// TwinCAT 3 PLC project PLC
// ProgramVersion: 3.1.4026.27
// libraries:
//   Tc2_Standard, * (Beckhoff Automation GmbH)
//   Tc2_System, * (Beckhoff Automation GmbH)
//   Tc3_EventLogger, * (Beckhoff Automation GmbH)
// project tree:
//   / PlcTask.TcTTO
//   POUs/ MAIN.TcPOU, FB_ActiveAlarmListener.TcPOU, I_ActiveAlarmList.TcIO, FB_Station.TcPOU, FB_StackLight.TcPOU
//   DUTs/ ST_EventListEntry.TcDUT
//   GVLs/ GVL_Params.TcGVL
// real-time tasks:
//   TASK PlcTask: cycle T#10ms, priority 20, ADS port 350

CONFIGURATION PLC
    RESOURCE PLC ON TwinCAT3
        TASK PlcTask(INTERVAL := T#10ms, PRIORITY := 20);
        PROGRAM MAIN WITH PlcTask : MAIN;
    END_RESOURCE
END_CONFIGURATION

// ---- DUTs/ST_EventListEntry.TcDUT
// One row of FB_ActiveAlarmListener (active alarm table and message ring buffer).
// Application independent: everything FB_TcEvent exposes, copied out of the callback.
TYPE ST_EventListEntry :
STRUCT
    bUsed       : BOOL;             // row in use = alarm is ACTIVE (raised, or cleared but waiting for confirmation)
    bIsAlarm    : BOOL;             // TRUE = alarm, FALSE = message
    bRaised     : BOOL;             // alarm state: TRUE = Raised, FALSE = cleared (row only kept while waiting for confirmation)
    eConfirmationState : TcEventConfirmationState;  // NotSupported / NotRequired / WaitForConfirmation / Confirmed / Reset
    nSequence   : UDINT;            // running number (messages only)
    eventClass  : GUID;             // event class
    nEventId    : UDINT;            // event id within the class
    eSeverity   : TcEventSeverity;  // Verbose..Critical
    nTimestamp  : ULINT;            // raise / send time stamped by the EventLogger, 100 ns since 1601-01-01 UTC
    nReceived   : ULINT;            // F_GetSystemTime when the listener callback ran (same clock, same unit)
    tLatency    : LTIME;            // nReceived - nTimestamp: raise -> visible in this table
    nSourceId   : UDINT;            // I_TcSourceInfo.nId   (application defined, e.g. station number)
    guidSource  : GUID;             // I_TcSourceInfo.guid
    sSourceName : STRING(255);      // I_TcSourceInfo.sName
END_STRUCT
END_TYPE

// ---- GVLs/GVL_Params.TcGVL
// Application (test harness) parameters.
{attribute 'qualified_only'}
VAR_GLOBAL CONSTANT
    cStations        : UDINT := 12;      // number of stations / stack lights
    cStationAlarms   : UDINT := 8;       // alarms per station (FB_Station.aAlarms, Event3..Event10)
END_VAR

// ---- POUs/I_ActiveAlarmList.TcIO
// Read-only view of an "active alarm list" + recent-message ring buffer.
//
// Consumers (stack lights, HMI summaries, interlocks, ...) depend on THIS, not on the
// FB that produces the list. FB_ActiveAlarmListener implements it from EventLogger
// callbacks; any other producer (e.g. a list built from the PLC's own FB_TcAlarm.bRaised
// states, or one fed by the .NET proxy over ADS) can implement it too and the consumers
// do not change.
//
// Alarm identity = event class + event id + source id.
// Rows are addressed 1..nMaxAlarms; GetAlarm is FALSE for an empty row.
// Messages are addressed by running sequence number 1..nMessageSequence; GetMessage is
// FALSE once a message has been overwritten in the ring buffer (size nMaxRecentMessages).
INTERFACE I_ActiveAlarmList EXTENDS __SYSTEM.IQueryInterface

// Number of raised alarms (any source) whose severity is within [eMinSeverity .. eMaxSeverity].
METHOD Count : UDINT
VAR_INPUT
    eMinSeverity : TcEventSeverity;
    eMaxSeverity : TcEventSeverity;
END_VAR
END_METHOD

// Number of raised alarms from source nSourceId (= FB_TcSourceInfo.nId the publisher used)
// whose severity is within [eMinSeverity .. eMaxSeverity].
METHOD CountBySource : UDINT
VAR_INPUT
    nSourceId    : UDINT;
    eMinSeverity : TcEventSeverity;
    eMaxSeverity : TcEventSeverity;
END_VAR
END_METHOD

// Number of raised alarms of one event class whose severity is within [eMinSeverity .. eMaxSeverity].
METHOD CountByEventClass : UDINT
VAR_INPUT
    eventClass   : GUID;
    eMinSeverity : TcEventSeverity;
    eMaxSeverity : TcEventSeverity;
END_VAR
END_METHOD

// TRUE if the alarm (event class + event id + source id) is currently raised.
METHOD IsActive : BOOL
VAR_INPUT
    eventClass : GUID;
    nEventId   : UDINT;
    nSourceId  : UDINT;
END_VAR
END_METHOD

// Copies row nIndex (1..nMaxAlarms) of the active alarm table. FALSE if the row is empty
// or nIndex is out of range. Iterate 1..nMaxAlarms to enumerate all raised alarms.
METHOD GetAlarm : BOOL
VAR_INPUT
    nIndex : UDINT;
END_VAR
VAR_IN_OUT
    stEntry : ST_EventListEntry;
END_VAR
END_METHOD

// Fetches the message with running number nSequence from the ring buffer.
// Returns FALSE if that message was never received or has already been overwritten.
// Typical use: remember nMessageSequence, then loop over the newer ones each cycle.
METHOD GetMessage : BOOL
VAR_INPUT
    nSequence : UDINT;
END_VAR
VAR_IN_OUT
    stEntry : ST_EventListEntry;
END_VAR
END_METHOD

// Number of alarms currently raised (rows in use).
PROPERTY nActiveAlarms : UDINT
GET
END_GET
END_PROPERTY

// Highest valid row index for GetAlarm.
PROPERTY nMaxAlarms : UDINT
GET
END_GET
END_PROPERTY

// Increments on every raise / clear / dispose. Compare to the last value seen to detect "list changed".
PROPERTY nAlarmChangeCounter : UDINT
GET
END_GET
END_PROPERTY

// Running number of the newest message received (0 = none yet).
PROPERTY nMessageSequence : UDINT
GET
END_GET
END_PROPERTY

// Ring buffer size: messages older than nMessageSequence - nMaxRecentMessages are gone.
PROPERTY nMaxRecentMessages : UDINT
GET
END_GET
END_PROPERTY

END_INTERFACE

// ---- POUs/MAIN.TcPOU
// Test harness: 12 stations publish events, ONE listener keeps the active alarm
// list and drives 12 stack lights - all in the PLC, no HMI involved.
//
// How to play (online, in the declaration part of MAIN):
//   1. set nTestStation (1..12) and nTestAlarm (1..8, see FB_Station header for the mapping)
//   2. pulse bTestRaise / bTestClear / bTestSendMessage
//   3. watch aActiveAlarms, aRecentMessages, aStackLights[n].bRed/bYellow/bGreen
PROGRAM MAIN
VAR
    aStations    : ARRAY[1..GVL_Params.cStations] OF FB_Station;      // event publishers (app specific)
    aStackLights : ARRAY[1..GVL_Params.cStations] OF FB_StackLight;   // decoder ring -> outputs (app specific)

    // the generic "active alarm list" (one per PLC) + the storage it works on (sized here, by the application)
    fbListener      : FB_ActiveAlarmListener;
    aActiveAlarms   : ARRAY[1..128] OF ST_EventListEntry;   // raised alarms
    aRecentMessages : ARRAY[1..32]  OF ST_EventListEntry;   // last 32 messages (ring buffer)
    fbFilter        : FB_TcEventFilter;
    bSubscribe   : BOOL := TRUE;
    hrSubscribe  : HRESULT;

    // --- test controls -------------------------------------------------------
    nTestStation       : UDINT := 1;   // 1..12
    nTestAlarm         : UDINT := 1;   // 1..8: 1,4,5 = Warning (yellow)  2,6,7 = Error (red)  3,8 = Critical (red)
    bTestRaise         : BOOL;         // raise aAlarms[nTestAlarm] on station nTestStation
    bTestClear         : BOOL;         // clear it again
    bTestSendMessage   : BOOL;         // green pulse
    bTestClearAll      : BOOL;         // clear every raised alarm on nTestStation
    hrTest             : HRESULT;

    // --- "noise" from another event class, to prove the filter ----------------
    // TC_EVENTS.MachineEvents is NOT in the listener's filter, so these must never
    // show up in fbListener even though they share source id 3 with station 3.
    fbMachineSource    : FB_TcSourceInfo;
    fbMachineMessage   : FB_TcMessage;
    fbMachineAlarm     : FB_TcAlarm;
    bMachineInit       : BOOL := TRUE;
    bTestMachineMessage    : BOOL;
    bTestMachineRaiseAlarm : BOOL;
    bTestMachineClearAlarm : BOOL;
    hrMachineTest      : HRESULT;

    // --- alarm WITH confirmation required: stays in the list after Clear(FALSE) until Confirm(); Clear(TRUE) ends it ---
    fbAckSource        : FB_TcSourceInfo;
    fbAckAlarm         : FB_TcAlarm;            // StationEvents.MotorFault, bWithConfirmation := TRUE, source id 13
    bAckInit           : BOOL := TRUE;
    bTestAckRaise      : BOOL;
    bTestAckConfirm    : BOOL;
    bTestAckClear      : BOOL;                  // Clear(FALSE): confirmation still required
    bTestAckClearReset : BOOL;                  // Clear(TRUE):  confirmation reset
    hrAckTest          : HRESULT;

    i : UDINT;
END_VAR

// 1) stations: give each its id and let it create its events (first cycle)
FOR i := 1 TO GVL_Params.cStations DO
    aStations[i].nStationId := i;
    aStations[i]();
END_FOR

// 2) subscribe the listener once - only to our station event class
IF bSubscribe THEN
    bSubscribe := FALSE;
    // TC_EVENTS.StationEvents is only a namespace; the class GUID is reachable through any of its
    // events (all carry the same uuidEventClass), so this matches ALL events of StationEvents.
    fbFilter.Clear().EventClass.EqualTo(TC_EVENTS.StationEvents.CycleComplete.uuidEventClass);
    hrSubscribe := fbListener.Subscribe2(fbFilter);
END_IF

// 3) process the event queue -> active alarm list (the FB body binds the arrays and runs Execute)
fbListener(aActiveAlarms := aActiveAlarms, aRecentMessages := aRecentMessages);

// 4) stack lights - each one filters the shared list by its own source id.
//    They see the listener only as I_ActiveAlarmList (fbListener is implicitly converted).
FOR i := 1 TO GVL_Params.cStations DO
    aStackLights[i](ipAlarmList := fbListener, nSourceId := i);
END_FOR

// 5) test controls
IF nTestStation >= 1 AND nTestStation <= GVL_Params.cStations THEN
    IF bTestSendMessage THEN bTestSendMessage := FALSE; hrTest := aStations[nTestStation].SendMessage();  END_IF
    IF bTestRaise       THEN bTestRaise       := FALSE; hrTest := aStations[nTestStation].Raise(nTestAlarm); END_IF
    IF bTestClear       THEN bTestClear       := FALSE; hrTest := aStations[nTestStation].Clear(nTestAlarm); END_IF
    IF bTestClearAll    THEN bTestClearAll    := FALSE; aStations[nTestStation].ClearAll();                  END_IF
END_IF

// 6) unrelated event class (filter test)
IF bMachineInit THEN
    bMachineInit := FALSE;
    fbMachineSource.Clear();
    fbMachineSource.nId   := 3;                 // deliberately collides with station 3
    fbMachineSource.sName := 'Machine';
    hrMachineTest := fbMachineMessage.CreateEx(TC_EVENTS.MachineEvents.MachineMessage, fbMachineSource);
    hrMachineTest := fbMachineAlarm.CreateEx(TC_EVENTS.MachineEvents.MachineAlarm, FALSE, fbMachineSource);
END_IF
IF bTestMachineMessage    THEN bTestMachineMessage    := FALSE; hrMachineTest := fbMachineMessage.Send(0);       END_IF
IF bTestMachineRaiseAlarm THEN bTestMachineRaiseAlarm := FALSE; hrMachineTest := fbMachineAlarm.Raise(0);        END_IF
IF bTestMachineClearAlarm THEN bTestMachineClearAlarm := FALSE; hrMachineTest := fbMachineAlarm.Clear(0, FALSE); END_IF

// 7) alarm with confirmation required (source id 13, no stack light; watch aActiveAlarms)
IF bAckInit THEN
    bAckInit := FALSE;
    fbAckSource.Clear();
    fbAckSource.nId   := 13;
    fbAckSource.sName := 'Ack test';
    hrAckTest := fbAckAlarm.CreateEx(TC_EVENTS.StationEvents.MotorFault, TRUE, fbAckSource);
END_IF
IF bTestAckRaise      THEN bTestAckRaise      := FALSE; hrAckTest := fbAckAlarm.Raise(0);        END_IF
IF bTestAckConfirm    THEN bTestAckConfirm    := FALSE; hrAckTest := fbAckAlarm.Confirm(0);      END_IF
IF bTestAckClear      THEN bTestAckClear      := FALSE; hrAckTest := fbAckAlarm.Clear(0, FALSE); END_IF
IF bTestAckClearReset THEN bTestAckClearReset := FALSE; hrAckTest := fbAckAlarm.Clear(0, TRUE);  END_IF

END_PROGRAM

// ---- POUs/FB_Station.TcPOU
// Reusable per-station event publisher.
// All events of a station share one FB_TcSourceInfo whose nId = station number and
// sName = 'Station n'. The listener uses nId to route the event to the right stack light.
//
// Event class TC_EVENTS.StationEvents (MyEvents.tmc), alarm index -> event:
//   message        CycleComplete   Info      'Cycle complete'
//   aAlarms[1]     MaintenanceDue  Warning   'Maintenance due'
//   aAlarms[2]     PartJam         Error     'Part jam'
//   aAlarms[3]     Overtemperature Critical  'Overtemperature'
//   aAlarms[4]     LowMaterial     Warning   'Low material'
//   aAlarms[5]     DoorOpen        Warning   'Door open'
//   aAlarms[6]     MotorFault      Error     'Motor fault'
//   aAlarms[7]     SensorFault     Error     'Sensor fault'
//   aAlarms[8]     EmergencyStop   Critical  'Emergency stop'
// Several alarms share a severity on purpose: the stack light must stay on until the
// LAST raised alarm of that severity is cleared.
FUNCTION_BLOCK FB_Station
VAR_INPUT
    nStationId : UDINT;     // 1..GVL_Params.cStations - set before the first call
END_VAR
VAR_OUTPUT
    bInitialized : BOOL;
    hrLastError  : HRESULT;                                        // last failed call (latched)
    aRaised      : ARRAY[1..GVL_Params.cStationAlarms] OF BOOL;    // live state of this station's own alarms
    nRaised      : UDINT;                                          // how many of them are raised
END_VAR
VAR
    fbSource   : FB_TcSourceInfo;
    fbMessage  : FB_TcMessage;
    aAlarms    : ARRAY[1..GVL_Params.cStationAlarms] OF FB_TcAlarm;
    aAlarmDefs : ARRAY[1..GVL_Params.cStationAlarms] OF TcEventEntry;
    hr         : HRESULT;
    i          : UDINT;
END_VAR

IF NOT bInitialized AND nStationId > 0 THEN
    bInitialized := TRUE;

    // source info = station identity (captured by the events at Create time)
    fbSource.Clear();
    fbSource.nId   := nStationId;
    fbSource.sName := CONCAT('Station ', UDINT_TO_STRING(nStationId));

    aAlarmDefs[1] := TC_EVENTS.StationEvents.MaintenanceDue;
    aAlarmDefs[2] := TC_EVENTS.StationEvents.PartJam;
    aAlarmDefs[3] := TC_EVENTS.StationEvents.Overtemperature;
    aAlarmDefs[4] := TC_EVENTS.StationEvents.LowMaterial;
    aAlarmDefs[5] := TC_EVENTS.StationEvents.DoorOpen;
    aAlarmDefs[6] := TC_EVENTS.StationEvents.MotorFault;
    aAlarmDefs[7] := TC_EVENTS.StationEvents.SensorFault;
    aAlarmDefs[8] := TC_EVENTS.StationEvents.EmergencyStop;

    hr := fbMessage.CreateEx(TC_EVENTS.StationEvents.CycleComplete, fbSource);
    IF FAILED(hr) THEN hrLastError := hr; END_IF
    FOR i := 1 TO GVL_Params.cStationAlarms DO
        hr := aAlarms[i].CreateEx(aAlarmDefs[i], FALSE, fbSource);
        IF FAILED(hr) THEN hrLastError := hr; END_IF
    END_FOR
END_IF

nRaised := 0;
FOR i := 1 TO GVL_Params.cStationAlarms DO
    aRaised[i] := aAlarms[i].bRaised;
    IF aRaised[i] THEN nRaised := nRaised + 1; END_IF
END_FOR

METHOD SendMessage : HRESULT
SendMessage := fbMessage.Send(0);
IF FAILED(SendMessage) THEN hrLastError := SendMessage; END_IF
END_METHOD

// Raises alarm nAlarm (1..GVL_Params.cStationAlarms, see table in the FB header).
METHOD Raise : HRESULT
VAR_INPUT
    nAlarm : UDINT;
END_VAR
IF nAlarm < 1 OR nAlarm > GVL_Params.cStationAlarms THEN
    Raise := DWORD_TO_DINT(16#80070057);  // E_INVALIDARG
ELSE
    Raise := aAlarms[nAlarm].Raise(0);
END_IF
IF FAILED(Raise) THEN hrLastError := Raise; END_IF
END_METHOD

// Clears alarm nAlarm (1..GVL_Params.cStationAlarms).
METHOD Clear : HRESULT
VAR_INPUT
    nAlarm : UDINT;
END_VAR
IF nAlarm < 1 OR nAlarm > GVL_Params.cStationAlarms THEN
    Clear := DWORD_TO_DINT(16#80070057);  // E_INVALIDARG
ELSE
    Clear := aAlarms[nAlarm].Clear(0, FALSE);
END_IF
IF FAILED(Clear) THEN hrLastError := Clear; END_IF
END_METHOD

// Clears every raised alarm of this station (test helper).
METHOD ClearAll
VAR
    n : UDINT;
END_VAR
FOR n := 1 TO GVL_Params.cStationAlarms DO
    IF aAlarms[n].bRaised THEN
        aAlarms[n].Clear(0, FALSE);
    END_IF
END_FOR
END_METHOD

END_FUNCTION_BLOCK

// ---- POUs/FB_StackLight.TcPOU
// APPLICATION SPECIFIC decoder ring: active alarm list -> one station's stack light.
// All knowledge about "stations" lives here; FB_ActiveAlarmListener knows nothing about them.
//   RED    flashes while any Error/Critical alarm from this source is raised
//   YELLOW flashes while any Warning (or lower) alarm from this source is raised
//   GREEN  flashes for 3 s after a message from this source
// The three colors are independent (a stack light can show more than one).
//
// Depends only on I_ActiveAlarmList, not on FB_ActiveAlarmListener: any list producer
// that implements the interface can drive it.
FUNCTION_BLOCK FB_StackLight
VAR_INPUT
    ipAlarmList   : I_ActiveAlarmList;      // the shared list (assign once; 0 = outputs stay off)
    nSourceId     : UDINT;                  // FB_TcSourceInfo.nId this station publishes with
END_VAR
VAR_OUTPUT
    bRed    : BOOL;
    bYellow : BOOL;
    bGreen  : BOOL;
    nActiveAlarms   : UDINT;                // diagnostics
    nActiveWarnings : UDINT;
    bMessageActive  : BOOL;
END_VAR
VAR
    bFirstCycle  : BOOL := TRUE;
    nLastMsgSeq  : UDINT;                   // last message sequence handled
    stMsg        : ST_EventListEntry;
    fbMsgTimer   : TON;
    fbBlinkTimer : TON;
    bBlink       : BOOL;
END_VAR
VAR CONSTANT
    tBlinkHalfPeriod : TIME := T#500MS;     // flash clock (1 Hz)
    tMsgFlashTime    : TIME := T#3S;        // how long GREEN flashes after a message
END_VAR

IF ipAlarmList = 0 THEN                     // no list connected -> everything off
    nActiveAlarms := 0; nActiveWarnings := 0; bMessageActive := FALSE;
    bRed := FALSE; bYellow := FALSE; bGreen := FALSE;
    RETURN;
END_IF

// --- alarms: just count rows of "my" source in the shared list ---
nActiveAlarms   := ipAlarmList.CountBySource(nSourceId, TcEventSeverity.Error,   TcEventSeverity.Critical);
nActiveWarnings := ipAlarmList.CountBySource(nSourceId, TcEventSeverity.Verbose, TcEventSeverity.Warning);

// --- messages: walk the ones that arrived since last cycle, react to "mine" ---
IF bFirstCycle THEN
    bFirstCycle := FALSE;
    nLastMsgSeq := ipAlarmList.nMessageSequence;
END_IF
IF ipAlarmList.nMessageSequence - nLastMsgSeq > ipAlarmList.nMaxRecentMessages THEN
    nLastMsgSeq := ipAlarmList.nMessageSequence - ipAlarmList.nMaxRecentMessages;  // ring buffer overrun
END_IF
WHILE nLastMsgSeq < ipAlarmList.nMessageSequence DO
    nLastMsgSeq := nLastMsgSeq + 1;
    IF ipAlarmList.GetMessage(nLastMsgSeq, stMsg) AND stMsg.nSourceId = nSourceId THEN
        bMessageActive := TRUE;
        fbMsgTimer(IN := FALSE);            // retrigger pulse
    END_IF
END_WHILE
fbMsgTimer(IN := bMessageActive, PT := tMsgFlashTime);
IF fbMsgTimer.Q THEN
    bMessageActive := FALSE;
END_IF

// --- flash clock ---
fbBlinkTimer(IN := NOT fbBlinkTimer.Q, PT := tBlinkHalfPeriod);
IF fbBlinkTimer.Q THEN
    bBlink := NOT bBlink;
END_IF

// --- decoder ring ---
bRed    := (nActiveAlarms   > 0) AND bBlink;
bYellow := (nActiveWarnings > 0) AND bBlink;
bGreen  :=  bMessageActive       AND bBlink;

END_FUNCTION_BLOCK

// ---- POUs/FB_ActiveAlarmListener.TcPOU
// Generic, application-independent "active alarm list" for the PLC.
// A PLC-side replacement for what FB_ReadTc3Events does for the visu event table,
// but without the visualization dependency and with structured data instead of text.
//
// Dependencies: Tc3_EventLogger, Tc2_System (MEMCMP), ST_EventListEntry, I_ActiveAlarmList.
//
// The APPLICATION owns the storage and passes it in as variable-length arrays (ARRAY[*]),
// so the table sizes are decided where the FB is used - no parameter list / GVL needed:
//   aActiveAlarms[]   - every alarm that is ACTIVE: raised, or cleared but still waiting for
//                       confirmation (same meaning as FB_TcAlarm.bActive). Added in OnAlarmRaised,
//                       removed when the alarm is neither raised nor waiting for confirmation
//                       (OnAlarmCleared / OnAlarmConfirmed / OnAlarmDisposed).
//   aRecentMessages[] - ring buffer of the last N messages, each tagged with a running nSequence
//
// Usage:
//   VAR
//       fbList          : FB_ActiveAlarmListener;
//       aActiveAlarms   : ARRAY[1..128] OF ST_EventListEntry;   // any size, any bounds
//       aRecentMessages : ARRAY[1..32]  OF ST_EventListEntry;
//   END_VAR
//   fbFilter.Clear().EventClass.EqualTo(<class>.uuidEventClass);        // or any other filter
//   fbList.Subscribe2(fbFilter);                                         // once; Subscribe() = everything
//   fbList(aActiveAlarms := aActiveAlarms, aRecentMessages := aRecentMessages);   // EVERY cycle
//   fbConsumer(ipAlarmList := fbList, ...);                              // consumers take I_ActiveAlarmList
//
// Notes:
//   - call the FB body every cycle: it binds the arrays and processes the event queue (callbacks below)
//   - only events raised AFTER Subscribe are seen (no history replay by the EventLogger)
//   - alarm identity = event class + event id + source id (what the EventLogger keys an alarm instance on)
//   - the fbEvent REFERENCE handed to the callbacks must not be stored, so fields are copied out
//   - I_ActiveAlarmList indexes rows 1..nMaxAlarms regardless of the array's declared bounds
FUNCTION_BLOCK FB_ActiveAlarmListener EXTENDS FB_ListenerBase2 IMPLEMENTS I_ActiveAlarmList
VAR_IN_OUT
    aActiveAlarms   : ARRAY[*] OF ST_EventListEntry;   // raised alarms (one row per alarm instance)
    aRecentMessages : ARRAY[*] OF ST_EventListEntry;   // message ring buffer
END_VAR
VAR_OUTPUT
    bTableOverflow  : BOOL;                            // an alarm could not be stored (latched, see Reset)
    hrLastError     : HRESULT;
    // Determinism check: the callbacks run inside this FB's body, in the PLC task. Latency from the
    // EventLogger's raise/send timestamp to the row being written is therefore bounded by the task
    // cycle (plus the publisher/listener call order within the cycle). Reset() clears tMaxLatency.
    tLastLatency    : LTIME;                           // of the most recent event (alarm or message)
    tMaxLatency     : LTIME;                           // worst case seen since start / Reset
    // callback counters (diagnostics)
    nRaisedCallbacks, nClearedCallbacks, nConfirmedCallbacks, nDisposedCallbacks, nMessageCallbacks : UDINT;
END_VAR
VAR
    // backing fields of the I_ActiveAlarmList properties
    _nActiveAlarms       : UDINT;   // rows in use in aActiveAlarms
    _nAlarmChangeCounter : UDINT;   // ++ on every raise / clear / dispose
    _nMessageSequence    : UDINT;   // ++ per received message
    stEmpty              : ST_EventListEntry;   // all zero, used to clear rows
    // IID of ITcAlarm (TcCOM interface behind every alarm event): lets the listener ask the
    // EventLogger for the alarm's raised / confirmation state inside the callback.
    // (plain VAR, not CONSTANT: TcQueryInterface takes the IID by reference)
    iidITcAlarm : IID := (Data1 := 16#EC6D4FF7, Data2 := 16#5805, Data3 := 16#4DDB,
                          Data4 := [16#A3, 16#16, 16#27, 16#89, 16#4E, 16#77, 16#D6, 16#44]);
END_VAR

// Binds the arrays (VAR_IN_OUT) and processes the EventLogger queue -> On... callbacks below.
hrLastError := SUPER^.Execute();

// Clears the active alarm table, the message ring buffer and the overflow flag.
// (Comparable to bClearTable of FB_ReadTc3Events.) Alarms raised later are picked up again.
METHOD Reset
VAR
    i : DINT;
END_VAR
FOR i := LOWER_BOUND(aActiveAlarms, 1) TO UPPER_BOUND(aActiveAlarms, 1) DO
    aActiveAlarms[i] := stEmpty;
END_FOR
FOR i := LOWER_BOUND(aRecentMessages, 1) TO UPPER_BOUND(aRecentMessages, 1) DO
    aRecentMessages[i] := stEmpty;
END_FOR
_nActiveAlarms  := 0;
bTableOverflow := FALSE;
tMaxLatency    := LTIME#0NS;
_nAlarmChangeCounter := _nAlarmChangeCounter + 1;
END_METHOD

// Number of raised alarms (any source) whose severity is within [eMinSeverity .. eMaxSeverity].
METHOD Count : UDINT
VAR_INPUT
    eMinSeverity : TcEventSeverity;
    eMaxSeverity : TcEventSeverity;
END_VAR
VAR
    i : DINT;
END_VAR
Count := 0;
FOR i := LOWER_BOUND(aActiveAlarms, 1) TO UPPER_BOUND(aActiveAlarms, 1) DO
    IF aActiveAlarms[i].bUsed
       AND aActiveAlarms[i].eSeverity >= eMinSeverity
       AND aActiveAlarms[i].eSeverity <= eMaxSeverity THEN
        Count := Count + 1;
    END_IF
END_FOR
END_METHOD

// Number of raised alarms from source nSourceId (= FB_TcSourceInfo.nId the publisher used)
// whose severity is within [eMinSeverity .. eMaxSeverity].
METHOD CountBySource : UDINT
VAR_INPUT
    nSourceId    : UDINT;
    eMinSeverity : TcEventSeverity;
    eMaxSeverity : TcEventSeverity;
END_VAR
VAR
    i : DINT;
END_VAR
CountBySource := 0;
FOR i := LOWER_BOUND(aActiveAlarms, 1) TO UPPER_BOUND(aActiveAlarms, 1) DO
    IF aActiveAlarms[i].bUsed
       AND aActiveAlarms[i].nSourceId = nSourceId
       AND aActiveAlarms[i].eSeverity >= eMinSeverity
       AND aActiveAlarms[i].eSeverity <= eMaxSeverity THEN
        CountBySource := CountBySource + 1;
    END_IF
END_FOR
END_METHOD

// Number of raised alarms of one event class whose severity is within [eMinSeverity .. eMaxSeverity].
METHOD CountByEventClass : UDINT
VAR_INPUT
    eventClass   : GUID;
    eMinSeverity : TcEventSeverity;
    eMaxSeverity : TcEventSeverity;
END_VAR
VAR
    i : DINT;
END_VAR
CountByEventClass := 0;
FOR i := LOWER_BOUND(aActiveAlarms, 1) TO UPPER_BOUND(aActiveAlarms, 1) DO
    IF aActiveAlarms[i].bUsed
       AND aActiveAlarms[i].eSeverity >= eMinSeverity
       AND aActiveAlarms[i].eSeverity <= eMaxSeverity
       AND MEMCMP(ADR(aActiveAlarms[i].eventClass), ADR(eventClass), SIZEOF(GUID)) = 0 THEN
        CountByEventClass := CountByEventClass + 1;
    END_IF
END_FOR
END_METHOD

// TRUE if the alarm (event class + event id + source id) is currently raised.
METHOD IsActive : BOOL
VAR_INPUT
    eventClass : GUID;
    nEventId   : UDINT;
    nSourceId  : UDINT;
END_VAR
IsActive := FindAlarm(eventClass, nEventId, nSourceId) >= LOWER_BOUND(aActiveAlarms, 1);
END_METHOD

// Copies row nIndex (1..nMaxAlarms) of the active alarm table. FALSE if the row is empty
// or nIndex is out of range. (1-based regardless of the array's declared bounds.)
METHOD GetAlarm : BOOL
VAR_INPUT
    nIndex : UDINT;
END_VAR
VAR_IN_OUT
    stEntry : ST_EventListEntry;
END_VAR
VAR
    i : DINT;
END_VAR
GetAlarm := FALSE;
IF nIndex >= 1 AND nIndex <= nMaxAlarms THEN
    i := LOWER_BOUND(aActiveAlarms, 1) + UDINT_TO_DINT(nIndex) - 1;
    IF aActiveAlarms[i].bUsed THEN
        stEntry  := aActiveAlarms[i];
        GetAlarm := TRUE;
    END_IF
END_IF
END_METHOD

// Fetches the message with running number nSequence from the ring buffer.
// Returns FALSE if that message was never received or has already been overwritten.
// Typical use: remember nMessageSequence, then loop over the newer ones each cycle.
METHOD GetMessage : BOOL
VAR_INPUT
    nSequence : UDINT;
END_VAR
VAR_IN_OUT
    stEntry : ST_EventListEntry;
END_VAR
VAR
    i : DINT;
END_VAR
GetMessage := FALSE;
IF nSequence = 0 OR nSequence > _nMessageSequence THEN
    RETURN;
END_IF
i := RingIndex(nSequence);
IF aRecentMessages[i].bUsed AND aRecentMessages[i].nSequence = nSequence THEN
    stEntry    := aRecentMessages[i];
    GetMessage := TRUE;
END_IF
END_METHOD

// Number of alarms currently raised (rows in use).
PROPERTY nActiveAlarms : UDINT
GET
nActiveAlarms := _nActiveAlarms;
END_GET
END_PROPERTY

// Highest valid row index for GetAlarm (= number of elements in aActiveAlarms).
PROPERTY nMaxAlarms : UDINT
GET
nMaxAlarms := DINT_TO_UDINT(UPPER_BOUND(aActiveAlarms, 1) - LOWER_BOUND(aActiveAlarms, 1) + 1);
END_GET
END_PROPERTY

// Increments on every raise / clear / dispose.
PROPERTY nAlarmChangeCounter : UDINT
GET
nAlarmChangeCounter := _nAlarmChangeCounter;
END_GET
END_PROPERTY

// Running number of the newest message received (0 = none yet).
PROPERTY nMessageSequence : UDINT
GET
nMessageSequence := _nMessageSequence;
END_GET
END_PROPERTY

// Ring buffer size (= number of elements in aRecentMessages).
PROPERTY nMaxRecentMessages : UDINT
GET
nMaxRecentMessages := DINT_TO_UDINT(UPPER_BOUND(aRecentMessages, 1) - LOWER_BOUND(aRecentMessages, 1) + 1);
END_GET
END_PROPERTY

// Array index in aRecentMessages for message sequence nSequence (>= 1).
METHOD PRIVATE RingIndex : DINT
VAR_INPUT
    nSequence : UDINT;
END_VAR
RingIndex := LOWER_BOUND(aRecentMessages, 1) + UDINT_TO_DINT((nSequence - 1) MOD nMaxRecentMessages);
END_METHOD

// Copies the fields of an incoming event into a table row and stamps the arrival time.
METHOD PRIVATE CopyEvent
VAR_INPUT
    fbEvent  : REFERENCE TO FB_TcEvent;
    bIsAlarm : BOOL;
END_VAR
VAR_IN_OUT
    stEntry : ST_EventListEntry;
END_VAR
VAR
    nNow : ULINT;
END_VAR
stEntry.bUsed      := TRUE;
stEntry.bIsAlarm   := bIsAlarm;
stEntry.eventClass := fbEvent.EventClass;
stEntry.nEventId   := fbEvent.nEventId;
stEntry.eSeverity  := fbEvent.eSeverity;
stEntry.nTimestamp := fbEvent.nTimestamp;

// raise -> here. Both stamps are Windows FILETIME (100 ns) from the same system clock.
nNow := F_GetSystemTime();
stEntry.nReceived := nNow;
IF nNow >= fbEvent.nTimestamp THEN
    stEntry.tLatency := ULINT_TO_LTIME((nNow - fbEvent.nTimestamp) * 100);
ELSE
    stEntry.tLatency := LTIME#0NS;
END_IF
tLastLatency := stEntry.tLatency;
IF stEntry.tLatency > tMaxLatency THEN
    tMaxLatency := stEntry.tLatency;
END_IF
IF fbEvent.ipSourceInfo <> 0 THEN
    stEntry.nSourceId   := fbEvent.ipSourceInfo.nId;
    stEntry.guidSource  := fbEvent.ipSourceInfo.guid;
    stEntry.sSourceName := fbEvent.ipSourceInfo.sName;
ELSE
    stEntry.nSourceId   := 0;
    stEntry.guidSource  := stEmpty.guidSource;
    stEntry.sSourceName := '';
END_IF
END_METHOD

// Array index of the alarm (class + id + source); LOWER_BOUND - 1 if not present.
METHOD PRIVATE FindAlarm : DINT
VAR_INPUT
    eventClass : GUID;
    nEventId   : UDINT;
    nSourceId  : UDINT;
END_VAR
VAR
    i : DINT;
END_VAR
FindAlarm := LOWER_BOUND(aActiveAlarms, 1) - 1;
FOR i := LOWER_BOUND(aActiveAlarms, 1) TO UPPER_BOUND(aActiveAlarms, 1) DO
    IF aActiveAlarms[i].bUsed
       AND aActiveAlarms[i].nEventId  = nEventId
       AND aActiveAlarms[i].nSourceId = nSourceId
       AND MEMCMP(ADR(aActiveAlarms[i].eventClass), ADR(eventClass), SIZEOF(GUID)) = 0 THEN
        FindAlarm := i;
        RETURN;
    END_IF
END_FOR
END_METHOD

// FindAlarm for an incoming event.
METHOD PRIVATE FindAlarmByEvent : DINT
VAR_INPUT
    fbEvent : REFERENCE TO FB_TcEvent;
END_VAR
VAR
    nSourceId : UDINT;
END_VAR
IF fbEvent.ipSourceInfo <> 0 THEN
    nSourceId := fbEvent.ipSourceInfo.nId;
END_IF
FindAlarmByEvent := FindAlarm(fbEvent.EventClass, fbEvent.nEventId, nSourceId);
END_METHOD

// Adds (or refreshes) a raised alarm in the table.
METHOD PRIVATE AddAlarm
VAR_INPUT
    fbEvent : REFERENCE TO FB_TcEvent;
END_VAR
VAR
    i, idx, nNone : DINT;
END_VAR
nNone := LOWER_BOUND(aActiveAlarms, 1) - 1;
idx   := FindAlarmByEvent(fbEvent);

IF idx = nNone THEN     // free slot
    FOR i := LOWER_BOUND(aActiveAlarms, 1) TO UPPER_BOUND(aActiveAlarms, 1) DO
        IF NOT aActiveAlarms[i].bUsed THEN
            idx := i;
            EXIT;
        END_IF
    END_FOR
END_IF

IF idx = nNone THEN
    bTableOverflow := TRUE;
    RETURN;
END_IF

IF NOT aActiveAlarms[idx].bUsed THEN
    _nActiveAlarms := _nActiveAlarms + 1;
END_IF
CopyEvent(fbEvent, TRUE, aActiveAlarms[idx]);
aActiveAlarms[idx].bRaised := TRUE;
QueryAlarmState(fbEvent, aActiveAlarms[idx]);
_nAlarmChangeCounter := _nAlarmChangeCounter + 1;
END_METHOD

// Asks the EventLogger for the alarm's current raised / confirmation state and stores it in the row.
// Returns FALSE if the event does not offer ITcAlarm (should not happen for alarm callbacks);
// the row then keeps bRaised as set by the caller and NotSupported as confirmation state.
METHOD PRIVATE QueryAlarmState : BOOL
VAR_INPUT
    fbEvent : REFERENCE TO FB_TcEvent;
END_VAR
VAR_IN_OUT
    stEntry : ST_EventListEntry;
END_VAR
VAR
    ipAlarm   : ITcAlarm;
    bIsRaised : BOOL32;
    eState    : TcEventConfirmationState;
END_VAR
QueryAlarmState := FALSE;
IF fbEvent.ipEvent = 0 THEN
    RETURN;
END_IF
IF SUCCEEDED(fbEvent.ipEvent.TcQueryInterface(iidITcAlarm, ADR(ipAlarm))) AND ipAlarm <> 0 THEN
    IF SUCCEEDED(ipAlarm.GetIsRaised(bIsRaised)) THEN
        stEntry.bRaised := bIsRaised <> 0;
    END_IF
    IF SUCCEEDED(ipAlarm.GetConfirmationState(eState)) THEN
        stEntry.eConfirmationState := eState;
    END_IF
    ipAlarm.TcRelease();
    QueryAlarmState := TRUE;
END_IF
END_METHOD

// Cleared / Confirmed callback: refresh the row's state and drop it once the alarm is
// neither raised nor waiting for confirmation (= FB_TcAlarm.bActive went FALSE).
METHOD PRIVATE UpdateAlarm
VAR_INPUT
    fbEvent    : REFERENCE TO FB_TcEvent;
    bConfirmed : BOOL;     // TRUE from OnAlarmConfirmed, FALSE from OnAlarmCleared
END_VAR
VAR
    idx : DINT;
END_VAR
idx := FindAlarmByEvent(fbEvent);
IF idx < LOWER_BOUND(aActiveAlarms, 1) THEN
    RETURN;                                   // not in the table (raised before Subscribe, or already removed)
END_IF

// best guess from the callback alone, then overwritten by the EventLogger's own answer if available
IF bConfirmed THEN
    aActiveAlarms[idx].eConfirmationState := TcEventConfirmationState.Confirmed;
ELSE
    aActiveAlarms[idx].bRaised := FALSE;
END_IF
QueryAlarmState(fbEvent, aActiveAlarms[idx]);

IF NOT aActiveAlarms[idx].bRaised
   AND aActiveAlarms[idx].eConfirmationState <> TcEventConfirmationState.WaitForConfirmation THEN
    RemoveAlarm(fbEvent);                     // inactive -> gone
ELSE
    _nAlarmChangeCounter := _nAlarmChangeCounter + 1;   // still active, state changed
END_IF
END_METHOD

// Removes an alarm from the table (no-op if not present).
METHOD PRIVATE RemoveAlarm
VAR_INPUT
    fbEvent : REFERENCE TO FB_TcEvent;
END_VAR
VAR
    idx : DINT;
END_VAR
idx := FindAlarmByEvent(fbEvent);
IF idx >= LOWER_BOUND(aActiveAlarms, 1) THEN
    aActiveAlarms[idx] := stEmpty;
    IF _nActiveAlarms > 0 THEN
        _nActiveAlarms := _nActiveAlarms - 1;
    END_IF
    _nAlarmChangeCounter := _nAlarmChangeCounter + 1;
END_IF
END_METHOD

METHOD OnAlarmRaised : HRESULT
VAR_INPUT
    fbEvent : REFERENCE TO FB_TcEvent;
END_VAR
nRaisedCallbacks := nRaisedCallbacks + 1;
AddAlarm(fbEvent);
OnAlarmRaised := S_OK;   // <> S_OK would pause further callbacks this cycle
END_METHOD

METHOD OnAlarmCleared : HRESULT
VAR_INPUT
    fbEvent : REFERENCE TO FB_TcEvent;
END_VAR
nClearedCallbacks := nClearedCallbacks + 1;
UpdateAlarm(fbEvent, FALSE);
OnAlarmCleared := S_OK;
END_METHOD

// Alarm instance released (FB_TcAlarm.Release / publisher stopped) - treat like cleared.
METHOD OnAlarmDisposed : HRESULT
VAR_INPUT
    fbEvent : REFERENCE TO FB_TcEvent;
END_VAR
nDisposedCallbacks := nDisposedCallbacks + 1;
RemoveAlarm(fbEvent);
OnAlarmDisposed := S_OK;
END_METHOD

// Confirm() on an alarm that was already cleared ends it -> row removed.
// Confirm() on a raised alarm only updates the confirmation state -> row stays.
METHOD OnAlarmConfirmed : HRESULT
VAR_INPUT
    fbEvent : REFERENCE TO FB_TcEvent;
END_VAR
nConfirmedCallbacks := nConfirmedCallbacks + 1;
UpdateAlarm(fbEvent, TRUE);
OnAlarmConfirmed := S_OK;
END_METHOD

// Messages are stateless: append to the ring buffer and bump the sequence.
METHOD OnMessageSent : HRESULT
VAR_INPUT
    fbEvent : REFERENCE TO FB_TcEvent;
END_VAR
VAR
    i : DINT;
END_VAR
nMessageCallbacks := nMessageCallbacks + 1;
_nMessageSequence := _nMessageSequence + 1;
i := RingIndex(_nMessageSequence);
CopyEvent(fbEvent, FALSE, aRecentMessages[i]);
aRecentMessages[i].nSequence := _nMessageSequence;
OnMessageSent := S_OK;
END_METHOD

END_FUNCTION_BLOCK
